FUNCTION_BLOCK A2X2_SPLIT_FWD_REV (* A2X2 passthrough (Socket zu Plug) plus 2 A2X Plugs, die den Vorwaerts- und den Rueckwaerts-Kanal spiegeln *)
  (* Standard: 61499-2; Function: IN -> OUT unveraendert, zusaetzlich an FWD_OUT gespiegelt. OUT -> IN (Rueckwaerts) unveraendert, zusaetzlich an REV_OUT gespiegelt.; Description: Copyright (c) 2026 HR Agrartechnik GmbH This program and the accompanying materials are made available under the terms of the Eclipse Public License 2.0 which is available at https://www.eclipse.org/legal/epl-2.0/ SPDX-License-Identifier: EPL-2.0 *)
  (* Version 1.0, 2026-11-13, Franz Höpfinger, HR Agrartechnik GmbH, Initial Version - Luecke in der Adapter-Familie geschlossen *)
  PACKAGE adapter::events::bidirectional;
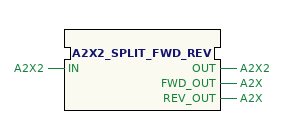
  SOCKETS
    IN : adapter::types::bidirectional::A2X2; (* bidirektionaler Eingang *)
  END_SOCKETS
  PLUGS
    OUT : adapter::types::bidirectional::A2X2; (* bidirektionaler Ausgang (Passthrough) *)
    FWD_OUT : adapter::types::unidirectional::A2X; (* spiegelt den Vorwaerts-Kanal (IN.EO* ) *)
    REV_OUT : adapter::types::unidirectional::A2X; (* spiegelt den Rueckwaerts-Kanal (OUT.EI* ) *)
  END_PLUGS
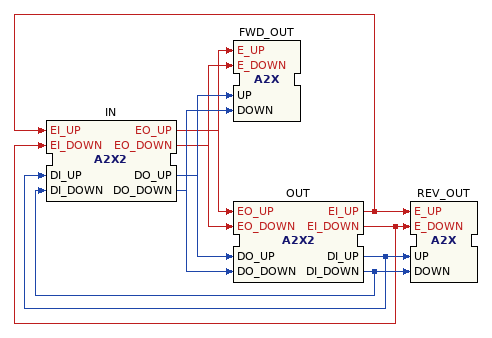
  EVENT_CONNECTIONS
    IN.EO_UP TO OUT.EO_UP;
    IN.EO_UP TO FWD_OUT.E_UP;
    OUT.EI_UP TO IN.EI_UP;
    OUT.EI_UP TO REV_OUT.E_UP;
    IN.EO_DOWN TO OUT.EO_DOWN;
    IN.EO_DOWN TO FWD_OUT.E_DOWN;
    OUT.EI_DOWN TO IN.EI_DOWN;
    OUT.EI_DOWN TO REV_OUT.E_DOWN;
  END_CONNECTIONS
  DATA_CONNECTIONS
    IN.DO_UP TO OUT.DO_UP;
    IN.DO_UP TO FWD_OUT.UP;
    OUT.DI_UP TO IN.DI_UP;
    OUT.DI_UP TO REV_OUT.UP;
    IN.DO_DOWN TO OUT.DO_DOWN;
    IN.DO_DOWN TO FWD_OUT.DOWN;
    OUT.DI_DOWN TO IN.DI_DOWN;
    OUT.DI_DOWN TO REV_OUT.DOWN;
  END_CONNECTIONS
END_FUNCTION_BLOCK
